(* PLC project g_timer_latch_mix, Anonymous Benchmark Suite 1.0 *)
(* stored: creationDateTime 2026-08-26T00:00:00 *)

PROGRAM g_timer_latch_mix
  VAR_INPUT
    Trig : BOOL;
    Ack : BOOL;
  END_VAR
  VAR_OUTPUT
    Alarm : BOOL;
  END_VAR
  VAR
    T0 : TON;
  END_VAR

(* LD diagram, written out as Structured Text *)
T0(IN := Trig, PT := T#30ms);
IF T0.Q THEN Alarm := TRUE; END_IF;
IF Ack THEN Alarm := FALSE; END_IF;
END_PROGRAM

CONFIGURATION Config0
  RESOURCE Res0 ON PLC
    TASK tcyclic(INTERVAL := T#10ms, PRIORITY := 0);
    PROGRAM inst0 WITH tcyclic : g_timer_latch_mix;
  END_RESOURCE
END_CONFIGURATION
